Fanuc KAREL source: KA00089.KL

PROGRAM KA00089
%NOLOCKGROUP
VAR
  SRC: JOINTPOS
  DST: POSITION
BEGIN
  DST = SRC
END KA00089
